Staubli VAL3: getLibName.pgx

public program getLibName(num& x_nLibNum, bool& x_bResult)
  local string l_sString
  local string l_sString1
  local num l_nPos
  local string l_sPath
  local num l_nlength
  local num l_nlength1
  local num l_nLength2
  local num l_nSize
  local string l_sTarget
  local num l_nLength
begin
  l_sPath=trajTemp:libPath()
  l_nlength=len("Disk://data/CustomerLib/lib")
  l_nlength1=len("/saveTRAJ/saveTRAJ.pjx")
  l_nLength2=len(l_sPath)
  l_nSize=l_nLength2-l_nlength1-l_nLength
  l_sTarget=mid(l_sPath,l_nSize,l_nlength)
  toNum(l_sTarget,x_nLibNum,x_bResult)
end
